Fanuc KAREL source: kd00022.KL

-- PROVISIONAL review KL for V770-1; original PC SHA256 bade85dbb53ad46e4fafa992b4ad4084ac237e870f0626797aacc3c2a77f04f0
-- Incomplete behavior may be omitted. Consult companion uncertainty JSON. Do not deploy.
PROGRAM KD00022
%NOLOCKGROUP
VAR
  I : INTEGER
  J : INTEGER
  B : BOOLEAN
  R : REAL
  S : STRING[80]
-- UNRESOLVED_DECL SAVED type=fd0010
BEGIN
  -- UNRESOLVED_PC offsets 5-12; opcodes 9D,23
  -- UNRESOLVED_PC offsets 17-21; opcodes 7F
END KD00022
